Fanuc KAREL source: kb00008.KL

-- PROVISIONAL review KL for V1013-1; original PC SHA256 36ef362ef83847e32c33ae7598bf1e8f7369683e1c614dfb13e94a5503eb6f05
-- Incomplete behavior may be omitted. Consult companion uncertainty JSON. Do not deploy.
PROGRAM KB00008
%NOLOCKGROUP
VAR
  P1 : REAL
  RESULT : REAL
BEGIN
  -- UNRESOLVED_PC offsets 5-16; opcodes 2E,23
  -- UNRESOLVED_PC offsets 21-36; opcodes 27,22,76,23
  -- UNRESOLVED_PC offsets 41-45; opcodes 7F
END KB00008
